Fanuc KAREL source: compact_preamble.KL

PROGRAM KD00022
%NOLOCKGROUP
VAR
I:INTEGER;J:INTEGER;B:BOOLEAN;R:REAL;S : STRING[80];SAVED:INTEGER
BEGIN
I=1
END KD00022
